// Application (test harness) parameters.
{attribute 'qualified_only'}
VAR_GLOBAL CONSTANT
    cStations        : UDINT := 12;      // number of stations / stack lights
    cStationAlarms   : UDINT := 8;       // alarms per station (FB_Station.aAlarms, Event3..Event10)
END_VAR

(* stored: Version 1.1.0.1
   GVL GVL_Params: Id {2d9dbeee-b719-44b5-a308-76f8862a66df} *)
